// Module : reçoit l'état agrégé de ses enfants, calculé par la station (docs/04 § 8)
INTERFACE I_Group

METHOD SetAggregate
VAR_INPUT
    eState : E_ObjState;
END_VAR
END_METHOD

END_INTERFACE

(* stored: Version 1.1.0.1, ProductVersion 3.1.4024.12
   Itf I_Group: Id {08e4e674-c993-5a6c-866f-0f47d17845a5}
   Method SetAggregate: Id {b3da1905-3fb9-58e4-b6df-e310336008da} *)
